// TwinCAT 3 PLC project MyLib
// Title: SampleLib
// Company: MyCompany
// ProjectVersion: 0.0.3
// ProgramVersion: 3.1.4026.25
// libraries:
//   Tc2_Standard, * (Beckhoff Automation GmbH)
//   Tc2_System, * (Beckhoff Automation GmbH)
// project tree:
//   POUs/ FB_Sum.TcPOU, FB_Diff.TcPOU, FB_Prod.TcPOU, FB_Div.TcPOU, FB_Mod.TcPOU
// real-time tasks:
//   TASK PlcTask: cycle T#10ms, priority 20, ADS port 350
//   TASK PlcTask1: cycle T#10ms, priority 21, ADS port 351

// ---- POUs/FB_Sum.TcPOU
// Function block for calculating the sum of two values
FUNCTION_BLOCK FB_Sum
VAR_INPUT
	var1: UINT;    // variable 1
	var2: UINT;    // variable 2
END_VAR
VAR_OUTPUT
	result : UINT; // result
END_VAR

// Calculation of the sum of two values; an error has been deliberately included in this example
result := var1 - var2;

END_FUNCTION_BLOCK

// ---- POUs/FB_Diff.TcPOU
// Function block for calculating the substraction of two values
FUNCTION_BLOCK FB_Diff
VAR_INPUT
	var1: UINT;    // variable 1
	var2: UINT;    // variable 2
END_VAR
VAR_OUTPUT
	result : UINT; // result
END_VAR

// Calculation of the substration of two values;
result := var1 - var2;

END_FUNCTION_BLOCK

// ---- POUs/FB_Prod.TcPOU
// Function block for calculating the product of two values
FUNCTION_BLOCK FB_Prod
VAR_INPUT
	var1: UINT;    // variable 1
	var2: UINT;    // variable 2
END_VAR
VAR_OUTPUT
	result : UINT; // result
END_VAR

// Calculation of the product of two values
result := var1 * var2;

END_FUNCTION_BLOCK

// ---- POUs/FB_Div.TcPOU
// Function block for calculating the division of two values
FUNCTION_BLOCK FB_Div
VAR_INPUT
	var1: UINT;    // variable 1
	var2: UINT;    // variable 2
END_VAR
VAR_OUTPUT
	result : UINT; // result
END_VAR

// Calculation of the division of two values
result := var1 / var2;

END_FUNCTION_BLOCK

// ---- POUs/FB_Mod.TcPOU
// Function block for calculating the modulo value of two variables
FUNCTION_BLOCK FB_Mod
VAR_INPUT
	var1: UINT;    // variable 1
	var2: UINT;    // variable 2
END_VAR
VAR_OUTPUT
	result : UINT; // result
END_VAR

// Calculation of the modulo value of two values
result := var1 Mod var2;

END_FUNCTION_BLOCK
